{region 'Documentation'}
(*!
<summary>Checks inequality with the forbidden ULINT value.</summary>
*)
{endregion}
FUNCTION_BLOCK AssertNotEqual_ULInt EXTENDS AssertionBase
VAR_INPUT
    IN : ULINT; //! Actual value checked or observed by this Assertion.
    Expected : ULINT; //! Value that must differ from IN under this Assertion's comparison rules.
END_VAR

SUPER^();

{region 'Documentation'}
(*!
<summary>Check inequality with the forbidden ULINT value.</summary>
*)
{endregion}
METHOD PROTECTED Assert
VAR
    Message : STRING(GVL_Constants.MessageLength);
    ExpectedText : STRING(GVL_Constants.AssertionValueLength);
    ActualText : STRING(GVL_Constants.AssertionValueLength);
END_VAR
IF NOT EvaluationActive THEN
    RETURN;
END_IF;

IF Result = E_Result.Error THEN
    RETURN;
END_IF;

IF Result = E_Result.Failed THEN
    RETURN;
END_IF;

IF IN = Expected THEN
    ExpectedText := ULINT_TO_STRING(Expected);
    ActualText := ULINT_TO_STRING(IN);
    Message := CONCAT('Assertion failed: values are equal but should differ. NotExpected = ',
        ExpectedText);
    Message := CONCAT(Message, ', Actual = ');
    Message := CONCAT(Message, ActualText);
    Message := CONCAT(Message, '.');
    Fail(Message := Message);
    RETURN;
END_IF;

Pass();
END_METHOD

END_FUNCTION_BLOCK

(* stored: Version 1.1.0.1
   POU AssertNotEqual_ULInt: Id {a5f5517d-369d-462e-8771-d94ba03c4c90}, SpecialFunc None
   Folder Internal: Id {a1e66d82-31b9-4df9-8f8e-f034748bb256}
   Method Assert: Id {ad773479-54b9-4bd0-8398-bce6dfa90a0c} *)
